(* PLC project Vn_mixed_big, Beckhoff Automation GmbH TwinCAT PLC Control 3.5.13.21 *)
(* stored: creationDateTime 1970-01-01T00:00:00 *)

PROGRAM Vn_mixed_big

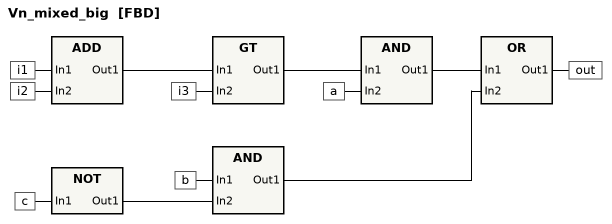
(* FBD diagram, written out as Structured Text *)
out := i1 + i2 > i3 AND a OR b AND NOT c;
END_PROGRAM
